// Mitsubishi GX Works2 project: Task_3   PLC: FX3G

PROGRAM MAIN
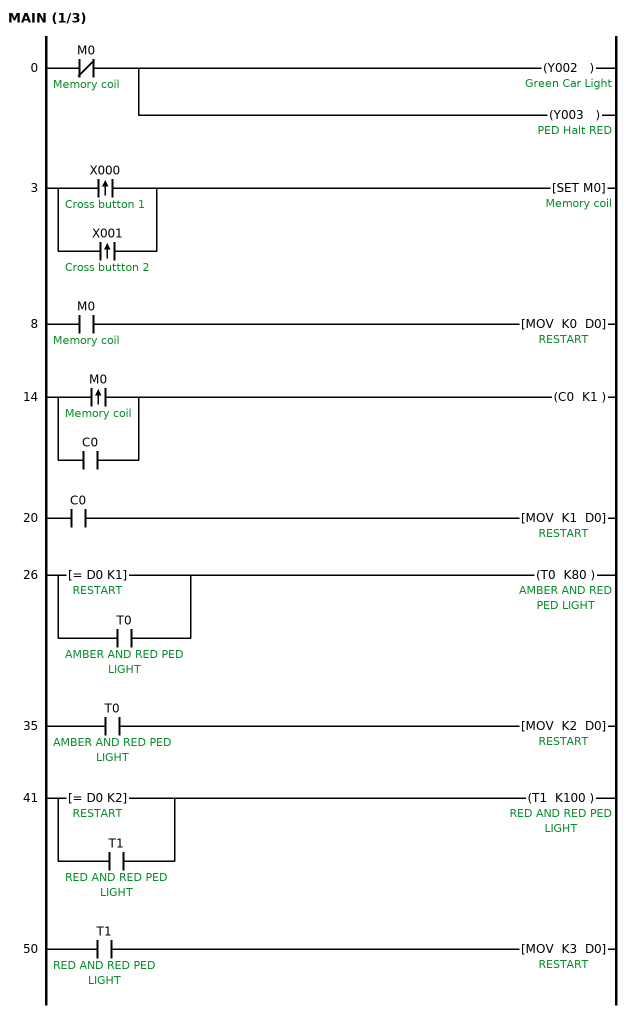
0     LDI     M0  ; Memory coil
      OUT     Y002  ; Green Car Light
      OUT     Y003  ; PED Halt RED
3     LDP     X000  ; Cross button 1
      ORP     X001  ; Cross buttton 2
      SET     M0  ; Memory coil
8     LD      M0  ; Memory coil
      MOV     K0 D0  ; RESTART
14    LDP     M0  ; Memory coil
      OR      C0
      OUT     C0 K1
20    LD      C0
      MOV     K1 D0
26    LD=     D0 K1  ; RESTART
      OR      T0  ; AMBER AND RED PED LIGHT
      OUT     T0 K80  ; AMBER AND RED PED LIGHT
35    LD      T0  ; AMBER AND RED PED LIGHT
      MOV     K2 D0
41    LD=     D0 K2  ; RESTART
      OR      T1  ; RED AND RED PED LIGHT
      OUT     T1 K100  ; RED AND RED PED LIGHT
50    LD      T1  ; RED AND RED PED LIGHT
      MOV     K3 D0
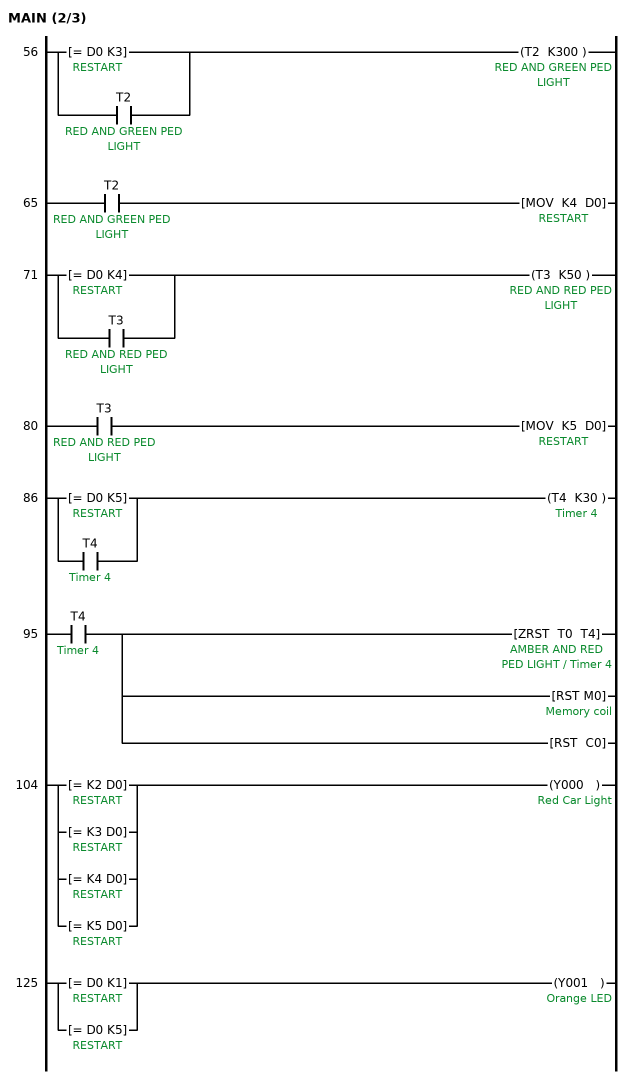
56    LD=     D0 K3  ; RESTART
      OR      T2  ; RED AND GREEN PED LIGHT
      OUT     T2 K300  ; RED AND GREEN PED LIGHT
65    LD      T2  ; RED AND GREEN PED LIGHT
      MOV     K4 D0
71    LD=     D0 K4  ; RESTART
      OR      T3  ; RED AND RED PED LIGHT
      OUT     T3 K50  ; RED AND RED PED LIGHT
80    LD      T3  ; RED AND RED PED LIGHT
      MOV     K5 D0
86    LD=     D0 K5  ; RESTART
      OR      T4  ; Timer 4
      OUT     T4 K30  ; Timer 4
95    LD      T4  ; Timer 4
      ZRST    T0 T4
      RST     M0  ; Memory coil
      RST     C0
104   LD=     K2 D0  ; RESTART
      OR=     K3 D0  ; RESTART
      OR=     K4 D0  ; RESTART
      OR=     K5 D0  ; RESTART
      OUT     Y000  ; Red Car Light
125   LD=     D0 K1  ; RESTART
      OR=     D0 K5  ; RESTART
      OUT     Y001  ; Orange LED
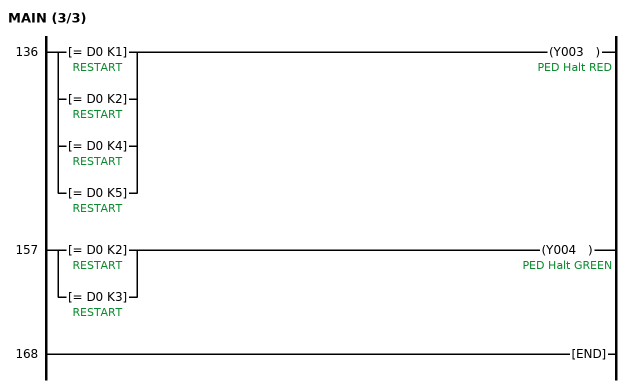
136   LD=     D0 K1  ; RESTART
      OR=     D0 K2  ; RESTART
      OR=     D0 K4  ; RESTART
      OR=     D0 K5  ; RESTART
      OUT     Y003  ; PED Halt RED
157   LD=     D0 K2  ; RESTART
      OR=     D0 K3  ; RESTART
      OUT     Y004  ; PED Halt GREEN
168   END
END_PROGRAM
